// TIA Portal V19 export
DATA_BLOCK "iFB_Control"   // DB21
// stored: InstanceOfName FB_Control, InstanceOfType FB
"FB_Control"
   // VAR_INPUT
   //    in_EmergencyStopHiPo : Bool;
   //    in_EmergencyStop : Bool;
   //    in_ResetButton : Bool;
   //    in_AutoSwitch : Bool;
   //    in_StartButton : Bool;
   //    in_StopButton : Bool;
   //    in_RobotTechMode : Bool;
   //    in_ServoIsOn : Bool;
   //    in_GateLocked : Bool;
   //    Blink : Bool;
   // END_VAR
   // VAR_OUTPUT
   //    ResetAlarms : Bool;
   //    ResetCycles : Bool;
   //    out_LedGreen : Bool;
   //    out_LedOrange : Bool;
   //    out_LedBlue : Bool;
   //    out_GateLock : Bool;
   //    out_GateLedStast : Bool;
   //    out_GateLedStop : Bool;
   //    out_RobotServoON : Bool;
   //    out_RobotExternalStart : Bool;
   //    out_RobotExternalHold : Bool;
   //    out_RobotAlarmReset : Bool;
   //    CurrentMachineState : Int;
   // END_VAR
   // VAR_IN_OUT
   //    EmergencyStop : Bool;
   //    ManualMode : Bool;
   //    AutoMode : Bool;
   //    AutoStarted : Bool;
   // END_VAR
   // VAR
   //    T_ResetAlarms { S7_SetPoint := 'True'} : TP_TIME;
   //    T_ResetCycles { S7_SetPoint := 'True'} : TON_TIME;
   // END_VAR
BEGIN
END_DATA_BLOCK
